// Mitsubishi GX Works2 project: 261012_기초회로_인터록회로_후입우선   PLC: Q03UDV

PROGRAM MAIN
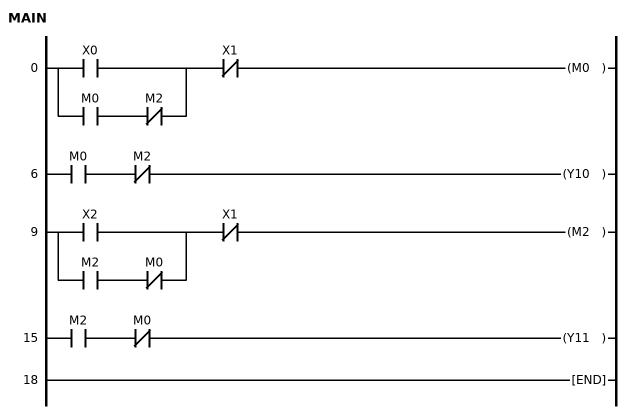
0     LD      X0
      LD      M0
      ANI     M2
      ORB
      ANI     X1
      OUT     M0
6     LD      M0
      ANI     M2
      OUT     Y10
9     LD      X2
      LD      M2
      ANI     M0
      ORB
      ANI     X1
      OUT     M2
15    LD      M2
      ANI     M0
      OUT     Y11
18    END
END_PROGRAM
